Fanuc KAREL source: KA00060.KL

PROGRAM KA00060
%NOLOCKGROUP
VAR
  SRC: POSITION
  DST: ARRAY[2] OF SHORT
BEGIN
  DST[1] = SRC
END KA00060
